(* IEC 61131-3 sources: openplc-editor-canopen/examples/canopen/scissor-lift/chassis-controller/pous/programs, 1 file *)

(* ---- main.st ---- *)
PROGRAM main
  VAR
    (* Inputs from the nodes, as the master maps them. *)
    platform_state AT %IB0 : USINT;
    joy_x AT %IW0 : INT;
    joy_y AT %IW1 : INT;
    estop_healthy AT platform_estop_healthy : BOOL;
    enable_switch AT platform_enable_switch : BOOL;
    drive_mode AT platform_drive_mode : BOOL;
    work_light AT platform_work_light : BOOL;
    valves_state AT %IB2 : USINT;
    lift_applied AT %IW2 : INT;
    drive_applied AT %IW3 : INT;
    supply_ok AT valves_supply_ok : BOOL;
    coil_fault AT valves_coil_fault : BOOL;
    sensor_state AT %IB4 : USINT;
    tilt AT %IW4 : INT;
    height AT %IW5 : UINT;
    load AT %IW6 : UINT;
    worklight_state AT %IB5 : USINT;
    (* Outputs to the nodes. *)
    lamp_ready AT platform_lamp_ready : BOOL;
    lamp_stop AT platform_lamp_stop : BOOL;
    lamp_tilt AT platform_lamp_tilt : BOOL;
    lamp_overload AT platform_lamp_overload : BOOL;
    lamp_warning AT platform_lamp_warning : BOOL;
    lamp_fault AT platform_lamp_fault : BOOL;
    lift_sp AT %QW0 : INT;
    drive_sp AT %QW1 : INT;
    valve_enable AT %QB1 : BYTE;
    light_cmd AT %QB2 : BYTE;
    display AT %QB3 : USINT;

    net : CANOPEN_NETWORK_STATE;
    light_node : CANOPEN_NODE_ENABLE;
    sensor_emcy : RECV_EMCY_DEV;
    valves_emcy : RECV_EMCY_DEV;
    isolate_valves : NMT;
    start_valves : NMT;
    read_serial : SDO_READ_STRING;
    read_seconds : SDO_READ4;
    write_ramp : SDO_WRITE4;
    poll : TON;

    estop, relay_off, neutral, need_neutral : BOOL;
    overload, valve_fault, isolated, tilt_alarm, base_ok, can_move, ready, lift_up_ok : BOOL;
    descent_hold, lowering : BOOL;
    want_seconds, want_ramp, serial_done : BOOL;
    last_mode, valves_were_up : BOOL;
    ramp_ms : UDINT;
    sensor_serial : STRING;
    operating_s : UDINT;
    stick : INT;
    raised, stowed : BOOL;
    last_height : UINT;
  END_VAR

(* The safety relay cuts the valves by itself; the program only sees its status and keeps the
   machine still until the stick has been in neutral after a reset. A node that is not operational
   reports nothing: that is a fault (the Fault lamp below), not an emergency stop. *)
base_ok := platform_state = OPERATIONAL AND (valves_state = OPERATIONAL OR isolated);
estop := platform_state = OPERATIONAL AND NOT estop_healthy;
relay_off := valves_state = OPERATIONAL AND NOT supply_ok;
neutral := ABS(joy_x) < 50 AND ABS(joy_y) < 50;
IF estop OR relay_off OR NOT base_ok THEN
  need_neutral := TRUE;
ELSIF neutral THEN
  need_neutral := FALSE;
END_IF;

(* The sensor's emergencies: overload on (3200h) and off (0000h). The valve module's coil fault is 5000h. *)
sensor_emcy(ENABLE := TRUE, DEVICE := sensor);
IF sensor_emcy.CONFIRM THEN
  IF sensor_emcy.EMCY.ERRORCODE = 16#3200 THEN
    overload := TRUE;
  ELSIF sensor_emcy.EMCY.ERRORCODE = 16#0000 THEN
    overload := FALSE;
  END_IF;
END_IF;
valves_emcy(ENABLE := TRUE, DEVICE := valves);
IF valves_emcy.CONFIRM THEN
  IF valves_emcy.EMCY.ERRORCODE = 16#5000 THEN
    valve_fault := TRUE;
  ELSIF valves_emcy.EMCY.ERRORCODE = 16#0000 THEN
    valve_fault := FALSE;
  END_IF;
END_IF;

(* A valve fault takes the valve module out of operation over NMT; pre-operational still sends
   emergencies. It is started again once the fault is cleared and the stick is in neutral. The state
   byte is the node's NMT state as it reports it: 127 is pre-operational. *)
isolate_valves(ENABLE := valve_fault AND valves_state = OPERATIONAL, DEVICE := valves, STATE := ENTER_PRE_OPERATIONAL);
IF valve_fault AND valves_state = OPERATIONAL THEN isolated := TRUE; END_IF;
start_valves(ENABLE := isolated AND NOT valve_fault AND neutral AND valves_state = 127,
             DEVICE := valves, STATE := START_REMOTE_NODE);
IF isolated AND valves_state = OPERATIONAL AND NOT valve_fault THEN isolated := FALSE; END_IF;

(* The platform floor is 1200 mm high when stowed; more than 300 mm above that counts as raised.
   A tilt of more than 3.00 degrees with the platform raised blocks lifting and driving, but the
   platform can still come down. The alarm ends within 2.50 degrees or when the platform is stowed. *)
raised := height > 1500;
stowed := height < 1260;
IF raised AND ABS(tilt) > 300 THEN
  tilt_alarm := TRUE;
ELSIF ABS(tilt) < 250 OR stowed THEN
  tilt_alarm := FALSE;
END_IF;

(* Moving needs the platform box and the valve module up, a healthy circuit, the enable switch and no fault. *)
net(ENABLE := TRUE);
can_move := base_ok AND NOT isolated AND NOT estop AND NOT relay_off AND NOT need_neutral AND enable_switch
            AND NOT valve_fault AND NOT coil_fault;
lift_up_ok := sensor_state = OPERATIONAL AND NOT overload AND NOT tilt_alarm;
stick := joy_y;
lowering := can_move AND NOT drive_mode AND stick < -50;

(* Descent stop: lowering through 2000 mm stops the platform. It goes on after the stick has been in
   neutral and is pushed down again, at no more than half speed below that height. *)
IF lowering AND last_height > 2000 AND height <= 2000 THEN descent_hold := TRUE; END_IF;
IF descent_hold AND neutral THEN descent_hold := FALSE; END_IF;
last_height := height;

lift_sp := 0;
drive_sp := 0;
valve_enable := 16#00;
IF can_move THEN
  valve_enable := 16#03;
  IF NOT drive_mode THEN
    IF stick > 0 AND lift_up_ok THEN
      lift_sp := stick;
    ELSIF stick < 0 AND NOT descent_hold THEN
      lift_sp := stick;
      IF height <= 2000 THEN lift_sp := MAX(stick, -500); END_IF;
    END_IF;
  ELSIF sensor_state = OPERATIONAL AND NOT tilt_alarm THEN
    (* Full speed when stowed, a fifth of it when raised. Steering is on and off, from the stick's side axis. *)
    IF raised THEN drive_sp := stick / 5; ELSE drive_sp := stick; END_IF;
    IF joy_x < -300 THEN valve_enable := valve_enable OR 16#04; END_IF;
    IF joy_x > 300 THEN valve_enable := valve_enable OR 16#08; END_IF;
  END_IF;
END_IF;

(* The lamps of the platform box. *)
ready := net.MANDATORY_UP AND base_ok AND sensor_state = OPERATIONAL AND NOT estop AND NOT relay_off
         AND NOT tilt_alarm AND NOT overload;
lamp_ready := ready;
lamp_stop := estop OR relay_off;
lamp_tilt := tilt_alarm;
lamp_overload := overload;
lamp_warning := tilt_alarm OR estop OR overload OR descent_hold;
lamp_fault := valve_fault OR coil_fault OR isolated OR NOT base_ok;

(* The display code: the first reason that keeps the machine still, else what it does. *)
IF estop THEN display := 1;
ELSIF relay_off THEN display := 2;
ELSIF NOT base_ok OR sensor_state <> OPERATIONAL THEN display := 9;
ELSIF valve_fault OR coil_fault OR isolated THEN display := 8;
ELSIF need_neutral AND NOT neutral THEN display := 4;
ELSIF descent_hold THEN display := 7;
ELSIF NOT enable_switch AND NOT neutral THEN display := 3;
ELSIF tilt_alarm AND (stick > 0 OR drive_mode) THEN display := 5;
ELSIF overload AND stick > 0 AND NOT drive_mode THEN display := 6;
ELSIF lift_sp > 0 THEN display := 10;
ELSIF lift_sp < 0 THEN display := 11;
ELSIF drive_sp <> 0 THEN display := 12;
ELSIF tilt_alarm THEN display := 5;
ELSIF overload THEN display := 6;
ELSE display := 0;
END_IF;

(* The optional work light node is on while the work light button is pressed. *)
light_node(ENABLE := TRUE, DEVICE := worklight, ACTIVE := work_light);
light_cmd := 16#00;
IF work_light AND worklight_state = OPERATIONAL THEN light_cmd := 16#01; END_IF;

(* The ramp-up time of the valve module depends on the mode: a gentle lift, a quicker drive. It is
   written when the mode changes and once each time the valve module comes up. *)
IF (drive_mode <> last_mode OR (valves_state = OPERATIONAL AND NOT valves_were_up)) AND NOT want_ramp THEN
  want_ramp := TRUE;
END_IF;
valves_were_up := valves_state = OPERATIONAL;
IF drive_mode THEN
  ramp_ms := 600;
ELSE
  ramp_ms := 1200;
END_IF;
write_ramp(ENABLE := want_ramp AND valves_state = OPERATIONAL, DEVICE := valves, INDEX := 16#2000, SUBINDEX := 4,
           DATA := UDINT_TO_DWORD(ramp_ms), DATALENGTH := 2);
IF write_ramp.CONFIRM OR write_ramp.ERROR <> 0 THEN
  want_ramp := FALSE;
  last_mode := drive_mode;
END_IF;

(* Once the sensor is up, read its serial number; every ten seconds read its operating time. *)
read_serial(ENABLE := sensor_state = OPERATIONAL AND NOT serial_done, DEVICE := sensor, INDEX := 16#2200, SUBINDEX := 1);
IF read_serial.CONFIRM THEN
  sensor_serial := read_serial.DATA;
  serial_done := TRUE;
END_IF;
poll(IN := NOT poll.Q, PT := T#10s);
IF poll.Q THEN
  want_seconds := TRUE;
END_IF;
read_seconds(ENABLE := want_seconds AND sensor_state = OPERATIONAL, DEVICE := sensor, INDEX := 16#2100, SUBINDEX := 4);
IF read_seconds.CONFIRM OR read_seconds.ERROR <> 0 THEN
  IF read_seconds.CONFIRM THEN
    operating_s := DWORD_TO_UDINT(read_seconds.DATA);
  END_IF;
  want_seconds := FALSE;
END_IF;

END_PROGRAM
